Fanuc KAREL source: kc00012.KL

PROGRAM KC00012
%STACKSIZE=65535
%PRIORITY=65535
%NOLOCKGROUP
VAR
I : INTEGER
J : INTEGER
K : INTEGER
R : REAL
B : BOOLEAN
S : STRING[80]
T : STRING[80]
AI : ARRAY[8] OF INTEGER
AB : ARRAY[244] OF BYTE
-- UNRESOLVED DECLARATIONS (source type spelling not recovered)
-- P : TYPE_0x001F (type_u16=0x001F)
-- Q : TYPE_0x001F (type_u16=0x001F)
-- QT : TYPE_0x1102 (type_u16=0x1102)
BEGIN
COPY_QUEUE(QT,AI,I,J,AI,K,I)
END KC00012
